FUNCTION_BLOCK "IPv4Parser"

VAR_INPUT
    ipText : STRING(254);
END_VAR

VAR_OUTPUT
    ipValue : UDINT;
END_VAR

BEGIN
    #ipValue := 0;
END_FUNCTION_BLOCK
